Staubli VAL3: safeTemp.pjx

--- safeTemp.pjx ---
Parameters version=s8.10.3Cs9_BS2093 stackSize=5000 millimeterUnit=true
Program file=start.pgx
Program file=stop.pgx
Data file=safeTemp.dtx
Type name=zoneItem path=Disk://source/template/zoneTemplate/zoneTemplate.pjx
Type name=sPoint path=Disk://source/template/sPointTemplate/sPointTemplate.pjx

--- safeTemp.dtx ---
public sPoint sSPoint
  [0]
    bool bActive
    pointRx pPointRx
    string sName
public zoneItem zZoneItem
  [0]
    pointRx pO
    pointRx pX
    pointRx pY
    frame fBase
    pointRx pFirst
    pointRx pSecond
    bool bActive
    string sID

--- start.pgx ---
program start()
begin
end

--- stop.pgx ---
program stop()
begin
end
